        IF Axis.StatusWord.3 OR NOT xEnable THEN
            iState := 999;
        ELSIF tonCapture.Q THEN
            // Trigger did not arrive within timeout
            tonCapture.IN := FALSE;
            iState := 999;
        ELSIF Axis.TouchProbe_StatusWord.1 THEN
            // Rising edge captured
            TouchProbe_Rising_Value       := Axis.TouchProbe_Rising_Value;
            Axis.TouchProbe_ControlWord.4 := FALSE;
            tonCapture.IN := FALSE;
            xDone_R := TRUE;
            iState := 40; // Hold result until xRisingCapture drops
        ELSIF NOT xExecute OR NOT Axis.TouchProbe_StatusWord.0 THEN
            Axis.TouchProbe_ControlWord.4 := FALSE;
            Axis.TouchProbe_ControlWord.5 := FALSE;
            tonCapture.IN := FALSE;
            iState := 0;
        END_IF

    30: // Wait for falling-edge trigger
        tonCapture(IN := TRUE,
                   PT := SEL(tCaptureTimeout = T#0S, tCaptureTimeout, T#999999S));

        IF Axis.StatusWord.3 OR NOT xEnable THEN
            iState := 999;
        ELSIF tonCapture.Q THEN
            tonCapture.IN := FALSE;
            iState := 999;
        ELSIF Axis.TouchProbe_StatusWord.2 THEN
            // Falling edge captured
            TouchProbe_Falling_Value      := Axis.TouchProbe_Falling_Value;
            Axis.TouchProbe_ControlWord.5 := FALSE;
            tonCapture.IN := FALSE;
            xDone_F := TRUE;
            iState := 50;
        ELSIF NOT xExecute OR NOT Axis.TouchProbe_StatusWord.0 THEN
            Axis.TouchProbe_ControlWord.4 := FALSE;
            Axis.TouchProbe_ControlWord.5 := FALSE;
            tonCapture.IN := FALSE;
            iState := 0;
        END_IF

    40: // Rising result hold - wait for application to drop xRisingCapture
        IF Axis.StatusWord.3 OR NOT xEnable THEN
            iState := 999;
        ELSIF NOT xRisingCapture THEN
            TouchProbe_Rising_Value := 0;
            xBusy := FALSE; xDone_R := FALSE;
            iState := 10;
        END_IF

    50: // Falling result hold - wait for application to drop xFallingCapture
        IF Axis.StatusWord.3 OR NOT xEnable THEN
            iState := 999;
        ELSIF NOT xFallingCapture THEN
            TouchProbe_Falling_Value := 0;
            xBusy := FALSE; xDone_F := FALSE;
            iState := 10;
        END_IF

    999:
        tonEnable.IN  := FALSE; tonCapture.IN := FALSE;
        tonEnable(PT := tEnableTimeout); tonCapture(PT := tCaptureTimeout);
        Axis.TouchProbe_ControlWord.4 := FALSE;
        Axis.TouchProbe_ControlWord.5 := FALSE;
        xBusy := FALSE; xError := TRUE;
        IF NOT xExecute OR xReset THEN
            xError := FALSE;
            iState := 0;
        END_IF

END_CASE

// -- Level A: unified progress projection (E_PROGRESS) --------------
IF    xError               THEN eProgress := PROGRESS_ERROR;
ELSIF xDone_R OR xDone_F    THEN eProgress := PROGRESS_DONE;   // at least one latch captured
ELSIF iState = 0            THEN eProgress := PROGRESS_INVALID;
ELSE                            eProgress := PROGRESS_BUSY;
END_IF

END_FUNCTION_BLOCK

// ---- POUs/FB_S7RTT_OTG.TcPOU
(* ============================================================
   FB_S7RTT_OTG - Online Trajectory Generator (OTG)
   SML v4 - Native implementation (replaces StruckigLight dependency)

   WHAT IT DOES:
   Generates a smooth, jerk-limited motion profile every PLC cycle.
   Given a target (position or velocity) and motion limits, it
   computes the next commanded position that respects:
     - MaxVelocity     [units/s]
     - MaxAcceleration [units/s^2]
     - MaxJerk         [units/s^3]

   TWO INTERFACES selected by ControlInterface:
   - FALSE (position): drive axis to TargetPosition; decelerate to
     stop at target without overshoot.
   - TRUE  (velocity): ramp to TargetVelocity; integrate to position.

   INITIALIZATION (v4 - explicit seed, fixes the fragile v3 auto-detect):
   In the mode-switch state, assert xInit = TRUE and write the actual
   axis position to CurrentPosition:
       otg.xInit           := TRUE;
       otg.CurrentPosition := DINT_TO_LREAL(Axis.Position_Actual_Value) / Scale;
   While xInit is TRUE the FB holds at CurrentPosition with zero velocity
   and acceleration.  In the motion loop call with xInit = FALSE.
   The v3 behaviour (re-init whenever CurrentPosition changed by value) was
   fragile: if the seed state lasted more than one cycle while the position
   moved, the OTG re-initialized every cycle and never advanced.  xInit makes
   the seed deterministic and decouples it from value comparison.

   ALGORITHM - S-curve (jerk-limited trapezoidal):
   Each cycle:
   1. Compute desired velocity:
      - Position mode: braking-limited velocity toward target
        v_brake = sqrt(2 * MaxAcceleration * |position_error|)
        (limits speed proportionally as target approaches - no overshoot)
      - Velocity mode: directly use TargetVelocity
   2. Compute desired acceleration = (v_desired - v_current) / dt
      Clamped to +/-MaxAcceleration
   3. Apply jerk limit: change in acceleration limited to MaxJerk * dt
   4. Integrate acceleration -> velocity (clamped to +/-MaxVelocity)
   5. Integrate velocity -> position
   6. Snap to target in position mode when within one-step distance

   NAMING NOTE:
   "CycleTIme" (capital I) is intentional - matches the typo present
   in the original OpenSML calls throughout the library.  Do not rename.
   All callers MUST use "CycleTIme :=" (v3 SyncPosition/SyncVelocity used the
   wrong "CycleTime" and did not compile - fixed in v4).

   COMPATIBILITY:
   Based on the StruckigLight FB_S7RTT_OTG.  v4 adds the xInit seed input,
   so callers must assert xInit during the seed cycle (see INITIALIZATION).
   ============================================================ *)

FUNCTION_BLOCK FB_S7RTT_OTG
VAR_INPUT
    ControlInterface : BOOL;    // FALSE = position interface, TRUE = velocity interface
    TargetPosition   : LREAL;   // Target position [user units] - used when ControlInterface=FALSE
    TargetVelocity   : LREAL;   // Target velocity [user units/s] - used when ControlInterface=TRUE
    CycleTIme        : LREAL;   // PLC task cycle time [s] - MUST match actual task period
    MaxVelocity      : LREAL;   // Velocity ceiling [user units/s] - must be > 0
    MaxAcceleration  : LREAL;   // Acceleration limit [user units/s^2] - must be > 0
    MaxJerk          : LREAL;   // Jerk limit [user units/s^3] - must be > 0
    // -- Seeding inputs ----------------------------------------
    // xInit: assert TRUE in the caller's mode-switch state to (re)seed the
    // integrator to CurrentPosition with zero velocity/acceleration.  Set FALSE
    // in the motion loop so the trajectory runs.  Deterministic - no value diff.
    xInit            : BOOL := FALSE;
    // CurrentPosition: actual axis position [user units], valid while xInit=TRUE.
    // Usage:  otg.CurrentPosition := DINT_TO_LREAL(Axis.Position_Actual_Value) / Scale;
    // Must be VAR_INPUT (not VAR) so CoDeSys allows external writes via dot notation.
    CurrentPosition  : LREAL := 0.0;
END_VAR
VAR_OUTPUT
    NewPosition : LREAL; // Commanded position for this cycle [user units]
    NewVelocity : LREAL; // Commanded velocity for this cycle [user units/s]
    xError      : BOOL;  // TRUE if inputs are invalid (zero limits or cycle time)
END_VAR
VAR
    // -- Internal integrator state -----------------------------
    _pos         : LREAL;   // Commanded position [user units]
    _vel         : LREAL;   // Commanded velocity [user units/s]
    _acc         : LREAL;   // Commanded acceleration [user units/s^2]

    // -- Initialization tracking -------------------------------
    _initialized : BOOL;    // FALSE until first seed is applied

    // -- Temporaries (declared here - no VAR_TEMP in FB) ------
    _desiredVel  : LREAL;
    _desiredAcc  : LREAL;
    _deltaAcc    : LREAL;
    _posError    : LREAL;
    _brakeVel    : LREAL;
    _snapDist    : LREAL;
END_VAR

// -- Input validation ------------------------------------------------------
IF CycleTIme <= 0.0 OR MaxVelocity <= 0.0 OR MaxAcceleration <= 0.0 THEN
    xError := TRUE;
    RETURN; // Outputs unchanged - caller must fix configuration
END_IF
xError := FALSE;

// If MaxJerk is zero or negative, disable jerk limiting by setting it very high
// (jerk limit is effectively infinite - pure trapezoidal profile)
IF MaxJerk <= 0.0 THEN MaxJerk := MaxAcceleration / CycleTIme; END_IF

// -- Explicit seed (v4) ----------------------------------------------------
// Caller asserts xInit=TRUE in its mode-switch state and writes CurrentPosition.
// While xInit is held (or until the first seed) the integrator is parked at the
// seed position with zero velocity/acceleration - deterministic, no value diff.
IF NOT _initialized OR xInit THEN
    _pos         := CurrentPosition;
    _vel         := 0.0; // Start from rest at seed position
    _acc         := 0.0;
    _initialized := TRUE;
    NewPosition  := _pos;
    NewVelocity  := _vel;
    RETURN; // Do not move on the initialization cycle
END_IF

// -- Step 1: Compute desired velocity --------------------------------------
IF NOT ControlInterface THEN

    // POSITION INTERFACE: compute braking-limited velocity toward target
    // v_brake = sqrt(2 * MaxAcceleration * |error|)
    // This is the maximum speed we can travel and still stop at the target
    // using MaxAcceleration. Staying within this speed prevents overshoot.
    _posError := TargetPosition - _pos;

    IF ABS(_posError) < 1.0E-10 THEN
        // Already at target (floating-point epsilon)
        _desiredVel := 0.0;
    ELSE
        // SQRT guard: argument must be >= 0 (ABS ensures this)
        _brakeVel   := SQRT(2.0 * MaxAcceleration * ABS(_posError));
        _brakeVel   := MIN(_brakeVel, MaxVelocity);

        // Apply direction: positive error -> positive velocity, negative -> negative
        IF _posError > 0.0 THEN
            _desiredVel := _brakeVel;
        ELSE
            _desiredVel := -_brakeVel;
        END_IF
    END_IF

ELSE

    // VELOCITY INTERFACE: ramp to requested velocity
    _desiredVel := TargetVelocity;

END_IF

// Clamp desired velocity to configured limits
_desiredVel := MAX(-MaxVelocity, MIN(MaxVelocity, _desiredVel));

// -- Step 2: Compute desired acceleration ----------------------------------
// Instantaneous acceleration needed to reach desired velocity in one step
// (before applying limits)
_desiredAcc := (_desiredVel - _vel) / CycleTIme;

// Clamp to MaxAcceleration
_desiredAcc := MAX(-MaxAcceleration, MIN(MaxAcceleration, _desiredAcc));

// -- Step 3: Apply jerk limit ----------------------------------------------
// Maximum change in acceleration per cycle = MaxJerk * dt
_deltaAcc := _desiredAcc - _acc;
_deltaAcc := MAX(-(MaxJerk * CycleTIme), MIN(MaxJerk * CycleTIme, _deltaAcc));
_acc := _acc + _deltaAcc;

// Re-clamp acceleration after jerk limiting (belt-and-suspenders)
_acc := MAX(-MaxAcceleration, MIN(MaxAcceleration, _acc));

// -- Step 4: Integrate acceleration -> velocity -----------------------------
_vel := _vel + _acc * CycleTIme;
_vel := MAX(-MaxVelocity, MIN(MaxVelocity, _vel));

// -- Step 5: Integrate velocity -> position --------------------------------
_pos := _pos + _vel * CycleTIme;

// -- Step 6: Snap to target in position mode --------------------------------
// When we are within one step distance of the target and velocity is small
// enough to stop within one cycle, snap to exact target to avoid steady-state
// oscillation around the target due to floating-point accumulation.
IF NOT ControlInterface THEN
    _snapDist := ABS(_vel) * CycleTIme; // Distance covered in one more cycle at current speed
    IF ABS(TargetPosition - _pos) <= _snapDist
       AND ABS(_vel) <= MaxAcceleration * CycleTIme THEN
        _pos := TargetPosition;
        _vel := 0.0;
        _acc := 0.0;
    END_IF
END_IF

// -- Outputs ---------------------------------------------------------------
NewPosition := _pos;
NewVelocity := _vel;

END_FUNCTION_BLOCK

// ---- POUs/FB_IoLink_In.TcPOU
(* ============================================================
   FB_IoLink_In - I/O bridge FB: INPUT image -> axis struct
   SML - I/O bridge (library FB)

   Copies DriveIn[] (the drive TxPDO image) into Axis[] (input
   fields), for all axes. Call at the START of the task, BEFORE the
   axis loop, so the computation uses fresh inputs (zero delay).

   Reusable: the arrays are passed by VAR_IN_OUT as ARRAY[*]
   (variable length) - no dependency on MAX_AXIS or on any
   application GVL. The application keeps the process image (e.g.
   GVL_IO.DriveIn) and its enable flag, and instantiates this FB.

   Precondition: DriveIn and Axis have the same bounds (one entry
   per axis). GATE: copies only when xEnable = TRUE.
   ============================================================ *)

FUNCTION_BLOCK FB_IoLink_In
VAR_INPUT
    xEnable : BOOL;   // TRUE = perform the copy; FALSE = bypass
END_VAR
VAR_IN_OUT
    DriveIn : ARRAY[*] OF ST_DriveIn;    // <- drive TxPDO image
    Axis    : ARRAY[*] OF OpenSML_Axis;  // -> axis struct (input fields written)
END_VAR
VAR
    i : DINT;
END_VAR

IF NOT xEnable THEN RETURN; END_IF

FOR i := LOWER_BOUND(Axis, 1) TO UPPER_BOUND(Axis, 1) DO
    Axis[i].StatusWord                   := DriveIn[i].StatusWord;
    Axis[i].Modes_of_operation_display   := DriveIn[i].Modes_of_operation_display;
    Axis[i].Torque_Actual_Value          := DriveIn[i].Torque_Actual_Value;
    Axis[i].Position_Actual_Value        := DriveIn[i].Position_Actual_Value;
    Axis[i].Velocity_Actual_Value        := DriveIn[i].Velocity_Actual_Value;
    Axis[i].Current_Actual_Value         := DriveIn[i].Current_Actual_Value;
    Axis[i].Following_Error_Actual_Value := DriveIn[i].Following_Error_Actual_Value;
    Axis[i].Error_Code                   := DriveIn[i].Error_Code;
    Axis[i].Digital_Inputs               := DriveIn[i].Digital_Inputs;
    Axis[i].TouchProbe_StatusWord        := DriveIn[i].TouchProbe_StatusWord;
    Axis[i].TouchProbe_Rising_Value      := DriveIn[i].TouchProbe_Rising_Value;
    Axis[i].TouchProbe_Falling_Value     := DriveIn[i].TouchProbe_Falling_Value;
END_FOR

END_FUNCTION_BLOCK

// ---- POUs/FB_IoLink_Out.TcPOU
(* ============================================================
   FB_IoLink_Out - I/O bridge FB: axis struct -> OUTPUT image
   SML - I/O bridge (library FB)

   Copies Axis[] (output fields) into DriveOut[] (the drive RxPDO
   image), for all axes. Call at the END of the task, AFTER the axis
   loop, so the outputs reflect the current cycle (zero delay).

   Reusable: the arrays are passed by VAR_IN_OUT as ARRAY[*]
   (variable length) - no dependency on MAX_AXIS or on any
   application GVL. The application keeps the process image (e.g.
   GVL_IO.DriveOut) and its enable flag, and instantiates this FB.

   Precondition: Axis and DriveOut have the same bounds (one entry
   per axis). GATE: copies only when xEnable = TRUE.
   ============================================================ *)

FUNCTION_BLOCK FB_IoLink_Out
VAR_INPUT
    xEnable : BOOL;   // TRUE = perform the copy; FALSE = bypass
END_VAR
VAR_IN_OUT
    Axis     : ARRAY[*] OF OpenSML_Axis;  // <- axis struct (output fields read)
    DriveOut : ARRAY[*] OF ST_DriveOut;   // -> drive RxPDO image
END_VAR
VAR
    i : DINT;
END_VAR

IF NOT xEnable THEN RETURN; END_IF

FOR i := LOWER_BOUND(Axis, 1) TO UPPER_BOUND(Axis, 1) DO
    DriveOut[i].ControlWord            := Axis[i].ControlWord;
    DriveOut[i].Modes_of_operation     := Axis[i].Modes_of_operation;
    DriveOut[i].Target_Position        := Axis[i].Target_Position;
    DriveOut[i].Profile_Velocity       := Axis[i].Profile_Velocity;
    DriveOut[i].Target_Velocity        := Axis[i].Target_Velocity;
    DriveOut[i].Target_Torque          := Axis[i].Target_Torque;
    DriveOut[i].Profile_Acceleration   := Axis[i].Profile_Acceleration;
    DriveOut[i].Profile_Deceleration   := Axis[i].Profile_Deceleration;
    DriveOut[i].Home_Offset            := Axis[i].Home_Offset;
    DriveOut[i].TouchProbe_ControlWord := Axis[i].TouchProbe_ControlWord;
END_FOR

END_FUNCTION_BLOCK

// ---- POUs/FB_Mapping_Out.TcPOU
(* ============================================================
   FB_Mapping_Out - MAPPING bridge FB: internal -> bus (state)
   SML - Level B / MAPPING (library FB)

   Copies the state/info from the internal structs into the bus
   UNIONs, for all axes:
     State[] -> StateBus[].stData   ,   Info[] -> InfoBus[].stData
   Call at the END of the task, after the axis loop.

   Reusable: arrays passed by VAR_IN_OUT as ARRAY[*] (variable
   length) - no dependency on MAX_AXIS or on any application GVL. The
   application keeps the bus UNION arrays (e.g. GVL_AXIS_MAP.State/Info)
   and its enable flag, and instantiates this FB.

   GATE: copies only when xEnable = TRUE.
   Runtime size check: if a struct exceeds its bus block (MAP_SIZE_STATE/INFO),
   the copy is blocked for safety (resize MAP_SIZE_* in GVL_SML_CONST).
   Precondition: all arrays have the same bounds (one entry per axis).
   ============================================================ *)

FUNCTION_BLOCK FB_Mapping_Out
VAR_INPUT
    xEnable : BOOL;   // TRUE = perform the copy; FALSE = bypass
END_VAR
VAR_IN_OUT
    State    : ARRAY[*] OF ST_AXIS_STATE;  // <- internal state
    Info     : ARRAY[*] OF ST_AXIS_INFO;   // <- internal info
    StateBus : ARRAY[*] OF U_AXIS_STATE;   // -> bus state (.stData)
    InfoBus  : ARRAY[*] OF U_AXIS_INFO;    // -> bus info  (.stData)
END_VAR
VAR
    i       : DINT;
    bSizeOk : BOOL;
END_VAR

IF NOT xEnable THEN RETURN; END_IF

// -- Bus block size check (safety) ----------------------------
bSizeOk := (SIZEOF(ST_AXIS_STATE) <= GVL_SML_CONST.MAP_SIZE_STATE)
       AND (SIZEOF(ST_AXIS_INFO)  <= GVL_SML_CONST.MAP_SIZE_INFO);
IF NOT bSizeOk THEN RETURN; END_IF   // blocked: resize MAP_SIZE_*

// -- Copy internal -> bus -------------------------------------
FOR i := LOWER_BOUND(State, 1) TO UPPER_BOUND(State, 1) DO
    StateBus[i].stData := State[i];
    InfoBus[i].stData  := Info[i];
END_FOR

END_FUNCTION_BLOCK

// ---- POUs/f_GetProgress.TcPOU
(* ============================================================
   f_GetProgress - Extracts the progress from a combined state
   SML v5 - Level A (new)

   eCombined = functional_state + E_PROGRESS  (progress band = 0..99)
   Returns only the progress part.

   Level B groundwork: not used by the Level A projection, provided
   as infrastructure for the combined state.
   ============================================================ *)

FUNCTION f_GetProgress : E_PROGRESS
VAR_INPUT
    eCombined : DINT;   // combined state = functional_state + progress
END_VAR

f_GetProgress := TO_INT(eCombined MOD GVL_SML_CONST.PROGRESS_SPAN);

END_FUNCTION

// ---- POUs/f_GetState.TcPOU
(* ============================================================
   f_GetState - Extracts the functional-state base from a combined state
   SML v5 - Level A (new)

   eCombined = functional_state + E_PROGRESS
   Returns functional_state (a multiple of PROGRESS_SPAN).
   In Level B the return type will become a dedicated enum
   (e.g. E_SML_AXIS_STATE).

   Level B groundwork: not used by the Level A projection.
   ============================================================ *)

FUNCTION f_GetState : DINT
VAR_INPUT
    eCombined : DINT;
END_VAR

f_GetState := (eCombined / GVL_SML_CONST.PROGRESS_SPAN) * GVL_SML_CONST.PROGRESS_SPAN;

END_FUNCTION
